// CFC twin of T_SafeRs_Tests: the same tests drawn as CFC diagrams, the way a TwinSAFE project is authored.
    FUNCTION_BLOCK T_SafeRs_Tests_CFC EXTENDS T_SafeCfcTestSuite
    VAR
    // Test_ResetDominantLatch
    group_1 : T_SafeGroup;
    fb_1 : T_SafeRs(group := group_1);
END_VAR

Test_ResetDominantLatch();

METHOD PRIVATE Test_ResetDominantLatch
// note: this text did not pass the execution check against the stored diagram
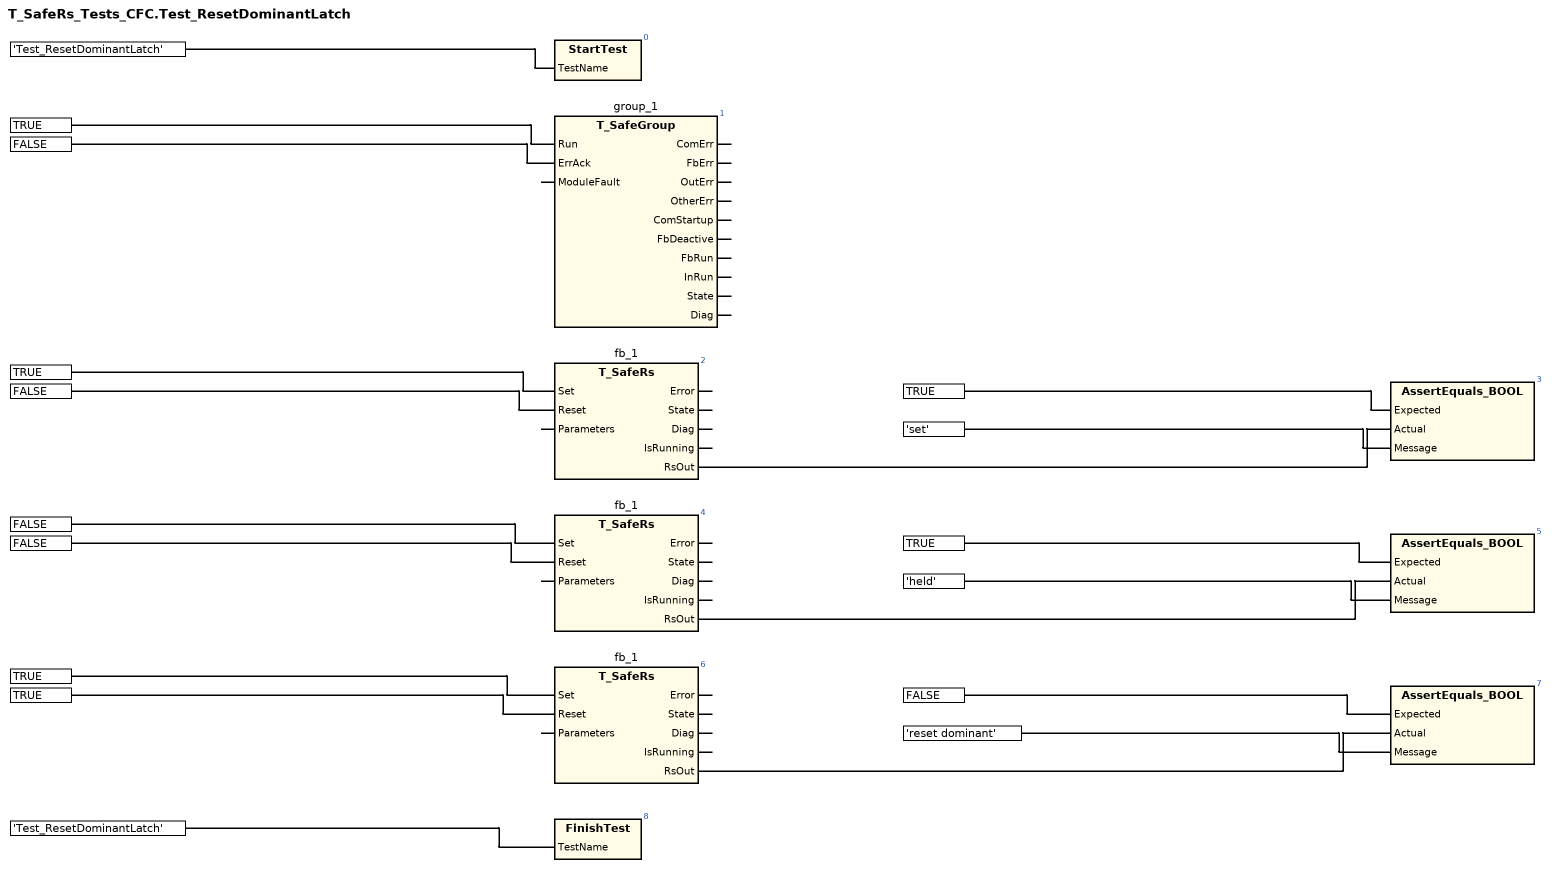
StartTest(TestName := 'Test_ResetDominantLatch');
group_1(Run := TRUE, ErrAck := FALSE); // T_SafeGroup
fb_1(Set := TRUE, Reset := FALSE); // T_SafeRs
AssertEquals_BOOL(Expected := TRUE, Actual := fb_1.RsOut, Message := 'set');
fb_1(Set := FALSE, Reset := FALSE); // T_SafeRs
AssertEquals_BOOL(Expected := TRUE, Actual := fb_1.RsOut, Message := 'held');
fb_1(Set := TRUE, Reset := TRUE); // T_SafeRs
AssertEquals_BOOL(Expected := FALSE, Actual := fb_1.RsOut, Message := 'reset dominant');
FinishTest(TestName := 'Test_ResetDominantLatch');
END_METHOD

END_FUNCTION_BLOCK

(* stored: Version 1.1.0.1, ProductVersion 3.1.4026.22
   POU T_SafeRs_Tests_CFC: Id {b4138d2a-3a49-5805-abd9-b74ddc966739}, SpecialFunc None
   Method Test_ResetDominantLatch: Id {011f9ec4-eca5-5e5b-aefd-8e908b32f92f} *)
